Fanuc KAREL source: kd00074.KL

PROGRAM KD00074
%STACKSIZE=65535
%PRIORITY=65535
%NOLOCKGROUP
VAR
I : INTEGER
J : INTEGER
B : BOOLEAN
R : REAL
S : STRING[80]
BEGIN
-- UNRESOLVED_PC line 10 opcodes [9C 3B] marker_code=0
END KD00074
